(* IEC 61131-3 sources: kns-pump-station/tests/POUs/Model/FB_HydraulicSolver_Test, 12 files *)

(* ---- FB_HydraulicSolver_Test.decl.st ---- *)
// Назначение: набор coUnit для FB_HydraulicSolver и F_PumpCurrent — законы подобия и рабочая точка насосов
//             на общий коллектор: один насос, параллельная работа, разные частоты и обратный клапан, напор ниже
//             статического, сухой ход, засор, осушенный приёмок, ток двигателя, давление PT201. Ожидаемые значения —
//             эталон tools_project/plant_reference.py (сценарии hydraulic.*), характеристика ST_PumpModelCfg по
//             умолчанию; допуски — REAL против float64 эталона.
// Автор:      kr0nsch
// Версия:     0.1.0
// Документ:   docs/DESIGN.md, разделы 11.3, 14.1
FUNCTION_BLOCK FB_HydraulicSolver_Test EXTENDS coUnit.FB_TestSuite
VAR CONSTANT
    R_LEVEL_M : REAL := 1.4;          // уровень подбора характеристики (DESIGN 11.3)
    R_EPS_Q : REAL := 0.005;          // допуск подачи, м³/ч
    R_EPS_H : REAL := 1.0E-3;         // допуск напора, м
    R_EPS_I : REAL := 1.0E-3;         // допуск тока, А
    R_EPS_P : REAL := 1.0E-4;         // допуск давления, бар
    R_UNDERLOAD_A : REAL := 12.0;     // порог недогрузки rUnderload_A (04 §10.3)
    R_IT_HH_A : REAL := 34.0;         // уставка HH IT1n1 (перечень)
    DW_NAN : DWORD := 16#7FC00000;
END_VAR

(* ---- AirLockZeroFlowLowCurrent.method.decl.st ---- *)
// Сухой ход насоса на 100 %: подача 0, ток 10,752 А — меньше порога недогрузки 12 А (PMI-15,
// DESIGN 11.3 ≈ 10,8 А).
METHOD PRIVATE AirLockZeroFlowLowCurrent
VAR
    fbDut : FB_HydraulicSolver; // проверяемый ФБ
    stCfg : ST_SimCfg;          // характеристика насоса по умолчанию (stCfg.stPump)
END_VAR

(* ---- ClogReducesFlowRaisesCurrent.method.decl.st ---- *)
// Засор на 100 %: подача 75,01 м³/ч (было 149,73), ток 34,299 А = 1,3 · 26,384 — выше HH 34 А
// (PMI-15, DESIGN 11.3 ≈ 34,3 А).
METHOD PRIVATE ClogReducesFlowRaisesCurrent
VAR
    fbDut : FB_HydraulicSolver; // проверяемый ФБ
    stCfg : ST_SimCfg;          // характеристика насоса по умолчанию (stCfg.stPump)
END_VAR

(* ---- ClogWithDryIntakeKeepsDryCurrent.method.decl.st ---- *)
// Засор при осушенном приёмке (0,25 м) и при сухом ходе насоса: подачи нет, ток — ток холостого хода
// 10,752 А, ниже порога недогрузки 12 А (DESIGN 11.2: «осушенный приёмок … ≈ 11 А, меньше порога 12 А»).
// Множитель засора к току без подачи не применяется — иначе 13,98 А маскировали бы сухой ход.
METHOD PRIVATE ClogWithDryIntakeKeepsDryCurrent
VAR
    fbDut : FB_HydraulicSolver; // проверяемый ФБ
    stCfg : ST_SimCfg;          // характеристика насоса по умолчанию (stCfg.stPump)
END_VAR

(* ---- DefaultsStoppedStaticHead.method.decl.st ---- *)
// Насосы стоят: подачи и токи 0, напор — статический Hgeo − h = 10,6 м, давление — столб за обратными
// клапанами ρ·g·Hgeo = 1,1772 бар.
METHOD PRIVATE DefaultsStoppedStaticHead
VAR
    fbDut : FB_HydraulicSolver; // проверяемый ФБ
    stCfg : ST_SimCfg;          // характеристика насоса по умолчанию (stCfg.stPump)
END_VAR

(* ---- IntakeDryNoFlow.method.decl.st ---- *)
// Осушенный приёмок (уровень 0,25 м < 0,30 м): насос на 100 % не подаёт, ток холостого хода 10,752 А,
// давление — столб 1,1772 бар.
METHOD PRIVATE IntakeDryNoFlow
VAR
    fbDut : FB_HydraulicSolver; // проверяемый ФБ
    stCfg : ST_SimCfg;          // характеристика насоса по умолчанию (stCfg.stPump)
END_VAR

(* ---- NoFlowBelowStaticHead.method.decl.st ---- *)
// 55 %: H0·s² = 10,44 м меньше статического напора 10,6 м — подачи нет, напор статический, ток
// холостого хода 5,011 А.
METHOD PRIVATE NoFlowBelowStaticHead
VAR
    fbDut : FB_HydraulicSolver; // проверяемый ФБ
    stCfg : ST_SimCfg;          // характеристика насоса по умолчанию (stCfg.stPump)
END_VAR

(* ---- NonFiniteSpeedTreatedAsStopped.method.decl.st ---- *)
// Неконечная скорость — насос не вращается: подача и ток 0, выходы конечны.
METHOD PRIVATE NonFiniteSpeedTreatedAsStopped
VAR
    fbDut : FB_HydraulicSolver; // проверяемый ФБ
    stCfg : ST_SimCfg;          // характеристика насоса по умолчанию (stCfg.stPump)
    uBits : PL.U_RealBits;
END_VAR

(* ---- ParallelPumpsMatchReference.method.decl.st ---- *)
// Параллельная работа: два по 75 % — 120,00 м³/ч (по 60,00); два по 100 % — 197,70; три по 100 % на
// 4,0 м — 224,17 м³/ч, напор 31,116 м (DESIGN 11.3, ASSUMPTIONS T9).
METHOD PRIVATE ParallelPumpsMatchReference
VAR
    fbDut : FB_HydraulicSolver; // проверяемый ФБ
    stCfg : ST_SimCfg;          // характеристика насоса по умолчанию (stCfg.stPump)
END_VAR

(* ---- PumpCurrentEdgeCases.method.decl.st ---- *)
// F_PumpCurrent: без вращения — 0; неконечный вход — 0; Pnom = 0 — 0; ток непрерывен при закрытии
// обратного клапана (подача 0,01 и 0 м³/ч дают одно значение 5,548 А на 60 %).
METHOD PRIVATE PumpCurrentEdgeCases
VAR
    stPump : ST_PumpModelCfg;   // характеристика по умолчанию
    uBits : PL.U_RealBits;
END_VAR

(* ---- SinglePumpMatchesReference.method.decl.st ---- *)
// Один насос: 100 % — 149,73 м³/ч, 20,913 м, 26,384 А, 2,1889 бар; 60 % — 41,32 м³/ч, 7,742 А,
// 1,2542 бар (DESIGN 11.3: 150 и 41 м³/ч; ASSUMPTIONS T8: ≈ 1,25 бар на минимуме).
METHOD PRIVATE SinglePumpMatchesReference
VAR
    fbDut : FB_HydraulicSolver; // проверяемый ФБ
    stCfg : ST_SimCfg;          // характеристика насоса по умолчанию (stCfg.stPump)
END_VAR

(* ---- UnequalSpeedsCheckValveClosed.method.decl.st ---- *)
// Разные частоты: 100 % и 60 % — у второго H0·0,36 = 12,4 м < напора 20,9 м, обратный клапан закрыт
// (подача 0, ток холостого хода 5,548 А); 100 % и 90 % — подают оба (120,46 и 60,77 м³/ч).
METHOD PRIVATE UnequalSpeedsCheckValveClosed
VAR
    fbDut : FB_HydraulicSolver; // проверяемый ФБ
    stCfg : ST_SimCfg;          // характеристика насоса по умолчанию (stCfg.stPump)
END_VAR
